TYPE "FRK_DeliveryResponse"
VERSION : 0.1
   STRUCT
      SchemaVersion : UInt;
      AckSequence : UDInt;
      Accepted : Bool;
   END_STRUCT;

END_TYPE

